Fanuc KAREL source: kx00026.compact.KL

PROGRAM KX00026
%STACKSIZE=65535
%PRIORITY=20
%NOLOCKGROUP
VAR
I : INTEGER
J : INTEGER
B : BOOLEAN
F : FILE
S : STRING[80]
P : XYZWPR
BEGIN
I=1
END KX00026
